Fanuc KAREL source: kb00166.compact.KL

PROGRAM KB00166
%STACKSIZE=65535
%PRIORITY=65535
%NOLOCKGROUP
%ENVIRONMENT REGOPE
VAR
P1 : INTEGER
P2 : JOINTPOS9
P3 : INTEGER
BEGIN
P1=1
P3=1
SET_JPOS_REG(P1,P2,P3,1)
END KB00166
